(* PLC project Vn_literal_assign, Beckhoff Automation GmbH TwinCAT PLC Control 3.5.13.21 *)
(* stored: creationDateTime 1970-01-01T00:00:00 *)

PROGRAM Vn_literal_assign

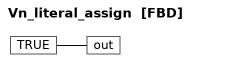
(* FBD diagram, written out as Structured Text *)
out := TRUE;
END_PROGRAM
